(* IEC 61131-3 sources: AyCD/PLC_Code (part 2) *)

            (* Outport: '<Root>/BRK_h_N1' *)
            BRK_h_N1 := b_BRK_h_N1;
            (* Outport: '<Root>/BRK_t_N1' *)
            BRK_t_N1 := b_BRK_t_N1;
            (* Outport: '<Root>/TLK' *)
            TLK := b_TLK;
            (* Outport: '<Root>/yc0_vec' *)
            FOR i := 0 TO 32 DO
                yc0_vec[i] := b_yc0_vec[i];
            END_FOR;
            (* End of Outport: '<Root>/yc0_vec' *)

            (* Outport: '<Root>/i_sel' *)
            i_sel := b_i_sel;
            (* Outport: '<Root>/vx_suave' *)
            vx_suave := b_vx_suave;
            (* Outport: '<Root>/vy_suave' *)
            vy_suave := b_vy_suave;
            (* Outport: '<Root>/recuperacion' *)
            recuperacion := b_recuperacion;
            (* Outport: '<Root>/modo_muerto' *)
            modo_muerto := b_modo_muerto;
            (* Outport: '<Root>/heartbeat' *)
            heartbeat := b_heartbeat;
            (* Outport: '<Root>/m_container' *)
            m_container := b_m_container;
            (* Outport: '<Root>/modo_auto' *)
            modo_auto := b_modo_auto;
            (* Outport: '<Root>/modo_manual' *)
            modo_manual := b_modo_manual;
            (* Outport: '<Root>/modo_manual_auto' *)
            modo_manual_auto := b_modo_manual_auto;
            (* Outport: '<Root>/modo_reposo' *)
            modo_reposo := b_modo_reposo;
            (* Outport: '<Root>/modo_error' *)
            modo_error := b_modo_error;
            (* Outport: '<Root>/sobrecarga' *)
            sobrecarga := b_sobrecarga;
        END_IF;
        IF plc_ts_counter1 >= 19 THEN
            plc_ts_counter1 := 0;
        ELSE
            plc_ts_counter1 := plc_ts_counter1 + 1;
        END_IF;
END_CASE;
END_FUNCTION_BLOCK
FUNCTION_BLOCK Suavizador_Cinematico
VAR_INPUT
    v_target: LREAL;
    v_act: LREAL;
    a_act: LREAL;
    A_MAX: LREAL;
    J_MAX: LREAL;
END_VAR
VAR_OUTPUT
    v_out: LREAL;
    a_out: LREAL;
END_VAR
VAR_TEMP
    err_v: LREAL;
    a_req: LREAL;
    jerk_req: LREAL;
    y: DINT;
    tmp: LREAL;
END_VAR
(* MATLAB Function 'Suavizador_Cinematico': '<S1>:334' *)
(* '<S1>:334:4' err_v = v_target - v_act; *)
err_v := v_target - v_act;
(* Error instantáneo de velocidad     *)
(* '<S1>:334:5' zona_lineal = 0.05; *)
(* Zona lineal cercana a cero para evitar singularidad en la raíz *)
(* Generación de aceleración deseada *)
(* '<S1>:334:8' if abs(err_v) < 1e-6 *)
tmp := ABS(err_v);
IF tmp < 1.0E-6 THEN
    (* Evita micro-oscilaciones cuando el error es prácticamente cero. *)
    (* '<S1>:334:9' v_out = v_target; *)
    v_out := v_target;
    (* '<S1>:334:10' a_out = 0; *)
    a_out := 0.0;
ELSE
    IF tmp > 0.05 THEN
        (* '<S1>:334:13' elseif abs(err_v) > zona_lineal *)
        (* '<S1>:334:14' a_req = sign(err_v) * sqrt(2 * J_MAX * abs(err_v)); *)
        IF err_v < 0.0 THEN
            y := -1;
        ELSIF err_v > 0.0 THEN
            y := 1;
        ELSE
            y := 0;
        END_IF;
        a_req := SQRT((2.0 * J_MAX) * tmp) * DINT_TO_LREAL(y);
        (* Región no lineal *)
    ELSE
        (* '<S1>:334:15' else *)
        (* '<S1>:334:16' a_req = (err_v / zona_lineal) * sqrt(2 * J_MAX * zona_lineal); *)
        a_req := SQRT((2.0 * J_MAX) * 0.05) * (err_v / 0.05);
        (* Región lineal cercana a cero para evitar pendiente infinita *)
    END_IF;
    (* Saturación de aceleración *)
    (* '<S1>:334:20' if a_req > A_MAX *)
    IF a_req > A_MAX THEN
        (* '<S1>:334:21' a_req = A_MAX; *)
        a_req := A_MAX;
    ELSIF a_req < ( -A_MAX) THEN
        (* '<S1>:334:22' elseif a_req < -A_MAX *)
        (* '<S1>:334:23' a_req = -A_MAX; *)
        a_req :=  -A_MAX;
    END_IF;
    (* Cálculo de jerk requerido *)
    (* '<S1>:334:27' jerk_req = (a_req - a_act) / 0.02; *)
    jerk_req := (a_req - a_act) / 0.02;
    (* Saturación de jerk *)
    (* '<S1>:334:29' if jerk_req > J_MAX *)
    IF jerk_req > J_MAX THEN
        (* '<S1>:334:30' jerk_req = J_MAX; *)
        jerk_req := J_MAX;
    ELSIF jerk_req < ( -J_MAX) THEN
        (* '<S1>:334:31' elseif jerk_req < -J_MAX *)
        (* '<S1>:334:32' jerk_req = -J_MAX; *)
        jerk_req :=  -J_MAX;
    END_IF;
    (* Integración discreta (Euler) *)
    (* '<S1>:334:36' a_out = a_act + jerk_req * 0.02; *)
    a_out := (jerk_req * 0.02) + a_act;
    (* '<S1>:334:37' v_out = v_act + a_out * 0.02; *)
    v_out := (a_out * 0.02) + v_act;
    (* Eliminación de deriva *)
    (* Forzar a cero absoluto si el joystick está suelto *)
    (* '<S1>:334:41' if abs(v_target) < 0.001 && abs(v_out) < 0.001 *)
    IF ABS(v_target) < 0.001 THEN
        IF ABS(v_out) < 0.001 THEN
            (* '<S1>:334:42' v_out = 0.0; *)
            v_out := 0.0;
            (* '<S1>:334:43' a_out = 0.0; *)
            a_out := 0.0;
        END_IF;
    END_IF;
END_IF;
END_FUNCTION_BLOCK
FUNCTION Check_Container: LREAL
VAR_INPUT
    i_pos: LREAL;
    y0_vec: ARRAY [0..32] OF LREAL;
END_VAR
VAR_TEMP
    temp1: BOOL;
END_VAR
(* MATLAB Function 'Check_Container': '<S1>:47' *)
(* '<S1>:47:4' if(i_pos<13 && y0_vec(i_pos)>0) *)
temp1 := FALSE;
IF i_pos < 13.0 THEN
    IF y0_vec[TRUNC(i_pos) - 1] > 0.0 THEN
        (* '<S1>:47:5' hay_container = 1; *)
        Check_Container := 1.0;
    ELSE
        temp1 := TRUE;
    END_IF;
ELSE
    temp1 := TRUE;
END_IF;
IF temp1 THEN
    IF (i_pos > 13.0) AND (i_pos < 33.0) THEN
        IF y0_vec[TRUNC(i_pos) - 1] > -18.0 THEN
            (* '<S1>:47:6' elseif(i_pos>13 && i_pos<33 && y0_vec(i_pos)>-18) *)
            (* '<S1>:47:7' hay_container = 1; *)
            Check_Container := 1.0;
        ELSE
            (* '<S1>:47:8' else *)
            (* '<S1>:47:9' hay_container = 0; *)
            Check_Container := 0.0;
        END_IF;
    ELSE
        (* '<S1>:47:8' else *)
        (* '<S1>:47:9' hay_container = 0; *)
        Check_Container := 0.0;
    END_IF;
END_IF;
END_FUNCTION
FUNCTION rt_floord: LREAL
VAR_INPUT
    u: LREAL;
END_VAR
rt_floord := DINT_TO_LREAL(TRUNC(u));
IF u = rt_floord THEN
    rt_floord := u;
ELSIF u < 0.0 THEN
    rt_floord := rt_floord - 1.0;
END_IF;
END_FUNCTION
FUNCTION_BLOCK isMember
VAR_INPUT
    a: LREAL;
END_VAR
VAR_OUTPUT
    tf: BOOL;
END_VAR
VAR
    b: ARRAY [0..2] OF SINT := 1,13,33;
END_VAR
VAR_TEMP
    k: DINT;
    exitg1: DINT;
END_VAR
tf := FALSE;
k := 0;
REPEAT
    exitg1 := 0;
    IF k < 3 THEN
        IF a = SINT_TO_LREAL(b[k]) THEN
            tf := TRUE;
            exitg1 := 1;
        ELSE
            k := k + 1;
        END_IF;
    ELSE
        exitg1 := 1;
    END_IF;
UNTIL NOT(exitg1 = 0)
END_REPEAT;
END_FUNCTION_BLOCK
FUNCTION_BLOCK PLC_CODER_TIMER
VAR_INPUT
    timerAction: INT;
    maxTime: DINT;
END_VAR
VAR_OUTPUT
    done: BOOL;
END_VAR
VAR
    plcTimer: TON;
    plcTimerExpired: BOOL;
END_VAR
CASE timerAction OF
    1:
        (* RESET *)
        plcTimer(IN:=FALSE, PT:=T#0ms);
        plcTimerExpired := FALSE;
        done := FALSE;
    2:
        (* AFTER *)
        IF (NOT(plcTimerExpired)) THEN
            plcTimer(IN:=TRUE, PT:=DINT_TO_TIME(maxTime));
        END_IF;
        plcTimerExpired := plcTimer.Q;
        done := plcTimerExpired;
    3:
        (* BEFORE *)
        IF (NOT(plcTimerExpired)) THEN
            plcTimer(IN:=TRUE, PT:=DINT_TO_TIME(maxTime));
        END_IF;
        plcTimerExpired := plcTimer.Q;
        done := NOT(plcTimerExpired);
END_CASE;
END_FUNCTION_BLOCK
VAR_GLOBAL CONSTANT
    Nivel_IN_NO_ACTIVE_CHILD: USINT := 0;
    Nivel_IN_Automata: USINT := 1;
    Nivel_IN_Muerto: USINT := 2;
    Nivel_IN_ABRIENDO_TLK: USINT := 1;
    Nivel_IN_CARGADO: USINT := 2;
    Nivel_IN_CERRANDO_TLK: USINT := 3;
    Nivel_IN_VACIO: USINT := 4;
    Nivel_IN_PULSOS_DOWN: USINT := 1;
    Nivel_IN_PULSOS_UP: USINT := 2;
    Nivel_IN_ERROR_FC_izq_der: USINT := 1;
    Nivel_IN_ERROR_FC_sup_inf: USINT := 2;
    Nivel_IN_ERROR_OTRO: USINT := 3;
    Nivel_IN_MANUAL: USINT := 4;
    Nivel_IN_MODO_AUTO: USINT := 5;
    Nivel_IN_RECUPERACION: USINT := 6;
    Nivel_IN_REPOSO: USINT := 7;
    Nivel_IN_AUTO_INIT: USINT := 1;
    Nivel_IN_MODO_MANUAL_SIMPLE: USINT := 2;
    Nivel_IN_MOVIMIENTO_CURVO: USINT := 3;
    c_Nivel_IN_MOVIMIENTO_CURVO: USINT := 4;
    c_Nivel_IN_SELECCION_TRAYEC: USINT := 5;
    Nivel_IN_SEL_DESTINO: USINT := 6;
    Nivel_IN_SEL_ORIGEN: USINT := 7;
    SS_INITIALIZE: SINT := 0;
    SS_STEP: SINT := 1;
END_VAR
VAR_GLOBAL
    plc_ts_counter1: DINT;
END_VAR
